# B&R Automation Studio project BrVideoPoker
Automation Studio 6.7.0.187; technology packages: mappServices 6.8.0, mappView 6.8.1, OpcUaCs 6.8.0

## Configuration Sim

CPU PC_any, AutomationRuntime D4.92, Build 11.3.0, Vc V4.72.5

### Task classes (Cpu.sw)
```
Cyclic#1:
  GameCode <- GameCode.prg
  UserSys <- UserSys.prg
  VisCtrl <- VisCtrl.prg
Binaries: arsvcreg, udbdef, TCData, arflatprv, arcoal, mvLoader, FWRules, Config_1, ashwac, User, sysconf, Config, asfw, arconfig, ashwd, Role, iomap
Libraries: PseudoRNG, AsIecCon, runtime, astime, AsIoTime, Cards, ArUser, arssl, ashw, arcert, fileio, sys_lib, aseth, dataobj, PokerHands, standard, MpUserX, MpBase
```

### Hardware
```
PC : PC_any v1.1.2.0 (OrderNumber=PC)
  ConfigurationID = BrVideoPoker_Sim
  FileDevice1
  FileDeviceName1 = USER
  FileDevicePath1 = USER_PATH
  ActivateOpcUa = 1
  OpcUa_SamplingTimer_Default = 4
  OpcUaInformationModels_PV_Version = 1
  ActivateFtpServer = 1
  ActivateWebServer = 1
  ActivateSdm = 1
```

### BRRole.brrole - PC/AccessAndSecurity/UserRoleSystem/BRRole.brrole
```
Element BR_Anonymous (Type=BRRole)
Element BR_Engineer (Type=BRRole)
Element BR_Observer (Type=BRRole)
Element BR_SafetyAdmin (Type=BRRole)
Element BR_SecurityAdmin (Type=BRRole)
```

- Physical/Sim/PC/IoMap.iom: same as Physical/Sim/PC/Cpu.per
- Physical/Sim/PC/PvMap.vvm: same as Physical/Sim/PC/Cpu.per
- Safety project (password-protected, skipped)

### Config.mpuserx - PC/mappServices/Config.mpuserx
```
Element UserMgmtX (Type=mpuserx)
  Mgr:
    AutoLogoutTime = 300
    UserNameLength = 3
    LoginAttempts = 5
  ServerSettings:
    Server:
      AdditionalUserData:
        [0] = mail
        [1] = telephoneNumber
  Groups:
    DefGroup#1:
      id = Administrators
      admin = TRUE
      rights:
        [0] = FullAccess
    DefGroup#2:
      id = Everyone
      level = 5
      admin = TRUE
```

### Config_1.mpuserxlogin - PC/mappServices/Config_1.mpuserxlogin
```
Element gUserXLogin (Type=mpuserxlogin)
```

## Configuration SuppC80

CPU 4PPC80.156B-13A, AutomationRuntime 6.8.1, Build 11.3.0

### Task classes (Cpu.sw)
```
Cyclic#1:
  GameCode <- GameCode.prg
  UserSys <- UserSys.prg
  VisCtrl <- VisCtrl.prg
Binaries: arsvcreg, udbdef, TCData, arflatprv, arcoal, mvLoader, FWRules, Config_1, ashwac, User, sysconf, Config, asfw, arconfig, ashwd, Role, iomap
Libraries: PseudoRNG, AsIecCon, runtime, astime, AsIoTime, Cards, ArUser, arssl, ashw, arcert, fileio, sys_lib, aseth, dataobj, PokerHands, standard, MpUserX, MpBase, AsBrStr
```

### Hardware
```
4PPC80_156B_13A : 4PPC80.156B-13A v1.4.0.0
  Connector IF2:
    AssignedOperatingSystem = ARemb
    ActivateDevice = 1
    ActivateSnmp = 2
  Connector IF3:
    OperatingSystem = ARemb
    ActivateDevice = 1
  Connector IF4:
    AssignedOperatingSystem = ARemb
  Connector IF5:
    AssignedOperatingSystem = GPOS
  Connector IF10:
    ActivateIna = 0
  ConfigurationID = BrVideoPoker_Sim
  Simulation = 1
  EnableDebugger = 1
  FileDevice1
  FileDeviceName1 = USER
  FileDevicePath1 = USER_PATH
  ActivateFtpServer = 1
  ActivateWebServer = 1
  ActivateSdm = 1
  LXTRemoteAccessUserWebGL = 
  LXTRemoteAccessPwdWebGL = 
```

- Physical/SuppC80/4PPC80_156B_13A/AccessAndSecurity/UserRoleSystem/BRRole.brrole: same as Physical/Sim/PC/AccessAndSecurity/UserRoleSystem/BRRole.brrole
- Physical/SuppC80/4PPC80_156B_13A/Cpu.per: same as Physical/Sim/PC/Cpu.per
- Physical/SuppC80/4PPC80_156B_13A/IoMap.iom: same as Physical/Sim/PC/Cpu.per
- Physical/SuppC80/4PPC80_156B_13A/PvMap.vvm: same as Physical/Sim/PC/Cpu.per
### Config.mpuserx - 4PPC80_156B_13A/mappServices/Config.mpuserx
```
Element UserMgmtX (Type=mpuserx)
  mapp.Gen:
    Audit = TRUE
  UserMgmtSystem:
    UserMgmtSystemType = 0
  ServerSettings:
    Server = ADServer
      Timeout = 10
      Mapping:
        TableName
      DisplayName = username
      AdditionalUserData:
        [0] = mail
        [1] = telephoneNumber
  PasswordPolicy:
    PasswordMaxAge = 0
    PasswordExpirationNotification = 0
    PasswordHistory = 0
    PasswordChangeReq = FALSE
    PasswordCase = TRUE
    PasswordAlpha = TRUE
    PasswordSpecial = TRUE
    PasswordLength = 8
  UserAccount:
    InvalidPasswordAttempts = 3
    UserExpirationTime = 0
    AutoLogoutTime = 3600
    UserNameLength = 1
    NoDelete = FALSE
    AdminUnlockTime = 3600
    EditSameLevel = 1
  ImportExport:
    ImportUser = 2
    ImportRole = 2
    ImportUnchecked = FALSE
    FileChecksum = 2
  Users:
    DefUser#1:
      id = Tester
      name
      lang
      measSystem = 0
  Roles:
    DefRole#1:
      id = Player
      level = 10
      admin = FALSE
```

- Physical/SuppC80/4PPC80_156B_13A/mappServices/Config_1.mpuserxlogin: same as Physical/Sim/PC/mappServices/Config_1.mpuserxlogin
## Logical view

Binary libraries used (declarations not repeated): operator, runtime, astime, AsIecCon, AsIoTime, ArUser, standard, MpUserX 6.8.0, MpBase 6.8.0, AsBrStr

### Global.typ - Global data types
```iecst
TYPE
	Player_typ : 	STRUCT
		Balance : REAL;
		Hand : ARRAY[0..4]OF Card_typ;
		HoldArr : ARRAY[0..4]OF BOOL;
		ChosenBet : REAL;
		Winnings : REAL;
		ActiveRound : BOOL;
		Result : FiveCardPoker_enum;
		LoggedIn : BOOL;
	END_STRUCT;
	Command_typ : 	STRUCT
		CMD_Confirm : BOOL;
		CMD_Action : BOOL;
	END_STRUCT;
END_TYPE
```

### Global.var - Global variables
```iecst
VAR
	gPlayer : Player_typ;
END_VAR
VAR CONSTANT
	BET_ARRAY : ARRAY[0..5] OF REAL := [0.1,0.2,0.5,1,2,5];
END_VAR
VAR
	gCurrentGame : GameVariant_enum;
	gCommand : Command_typ;
	gPayTable : PayTable_typ;
	gDeck : DeckFB;
	gPasswordInput : STRING[24];
	gUsernameInput : STRING[80];
END_VAR
```

### Package Logical/Libraries - Global libraries

### Library Logical/Libraries/Cards (IEC)

#### Types.typ - Exported data types
```iecst
TYPE
	Faces_enum :
		(
		CARD_TWO,
		CARD_THREE,
		CARD_FOUR,
		CARD_FIVE,
		CARD_SIX,
		CARD_SEVEN,
		CARD_EIGHT,
		CARD_NINE,
		CARD_TEN,
		CARD_JACK,
		CARD_QUEEN,
		CARD_KING,
		CARD_ACE
		);
	Suits_enum :
		(
		SUIT_HEARTS,
		SUIT_CLUBS,
		SUIT_DIAMONDS,
		SUIT_SPADES
		);
	Card_typ : 	STRUCT
		Face : Faces_enum;
		Suit : Suits_enum;
	END_STRUCT;
	DeckState :
		(
		DECKSTATE_INIT,
		DECKSTATE_IDLE,
		DECKSTATE_SHUFFLE,
		DECKSTATE_ERROR
		);
END_TYPE
```

#### Cards.fun - Exported functions and function blocks
```iecst
{REDUND_ERROR} FUNCTION SwapCard : BOOL (*Swap the place of two cards within deck*) (*$GROUP=User,$CAT=User,$GROUPICON=User.png,$CATICON=User.png*)
	VAR_INPUT
		Deck : REFERENCE TO ARRAY[0..51] OF Card_typ;
		CardIndexA : USINT;
		CardIndexB : USINT;
	END_VAR
	VAR
		TempCard : Card_typ;
	END_VAR
END_FUNCTION

FUNCTION_BLOCK DeckFB (*Core funciton block of the library*)
	VAR_INPUT
		CMD_Shuffle : BOOL;
		Enable : BOOL;
	END_VAR
	VAR_OUTPUT
		Deck : ARRAY[0..51] OF Card_typ;
		Active : BOOL;
		CommandDone : BOOL;
	END_VAR
	VAR
		IndexI : USINT;
		IndexJ : USINT;
		IndexR : USINT;
		ShuffleCount : USINT := 5;
		FaceIndex : USINT;
		SuitIndex : USINT;
		State : DeckState;
		Initialized : BOOL;
		Randy : PRNG;
	END_VAR
END_FUNCTION_BLOCK
```

#### CardsFB.st
```iecst
(* Deck Funtionality *)
FUNCTION_BLOCK DeckFB
	CASE State OF
		DECKSTATE_INIT:
			IF Enable AND NOT Initialized THEN
				//Initialize unshuffled deck
				FOR SuitIndex := 0 TO 3 DO
					FOR FaceIndex := 0 TO 12 DO
						Deck[SuitIndex*13+FaceIndex].Face := FaceIndex;
						Deck[SuitIndex*13+FaceIndex].Suit := SuitIndex;
					END_FOR;
				END_FOR;

				//Initialize RNG
				Randy(Multiplier := 4, Increment := 13, Seed := AsIOTimeStamp());

				State := DECKSTATE_IDLE;
				Active := TRUE;
				Initialized := TRUE;
			END_IF

		DECKSTATE_IDLE:
			IF CommandDone AND CMD_Shuffle THEN
				CommandDone := FALSE;
				CMD_Shuffle := FALSE;
			END_IF

			IF CMD_Shuffle THEN
				State := DECKSTATE_SHUFFLE;
			END_IF

		DECKSTATE_SHUFFLE:
			FOR IndexI := 0 TO ShuffleCount DO
				FOR IndexJ := 0 TO 51 DO
					Randy.CMD_Generate := TRUE;
					Randy();

					IndexR := UDINT_TO_USINT(  IndexJ + (Randy.Result MOD (52-IndexJ)));
					SwapCard(ADR(Deck), IndexJ, IndexR);
				END_FOR;
			END_FOR;

			CommandDone := TRUE;
			State := DECKSTATE_IDLE;

		DECKSTATE_ERROR:

	END_CASE;

END_FUNCTION_BLOCK
```

#### SwapCard.st
```iecst
(* Swap the place of two cards within deck *)
FUNCTION SwapCard
	TempCard := Deck[CardIndexA];
	Deck[CardIndexA] := Deck[CardIndexB];
	Deck[CardIndexB] := TempCard;
END_FUNCTION
```

### Library Logical/Libraries/PseudoRNG (IEC, version 1.00.1) - This library generates pseudo random numbers.

#### Constants.var - Exported constants
```iecst
VAR CONSTANT
	RAND_MAX : UINT := 32797; (*Maximum possible value for random number.*)
END_VAR
```

#### PseudoRNG.fun - Exported functions and function blocks
```iecst
FUNCTION_BLOCK PRNG
	VAR_INPUT
		Multiplier : {REDUND_UNREPLICABLE} UINT := 16; (*Multiplier parameter in formula*)
		Increment : {REDUND_UNREPLICABLE} UINT := 0; (*Increment parameter in formula*)
		CMD_Generate : {REDUND_UNREPLICABLE} BOOL; (*Input used to trigger generation*)
		Seed : UDINT; (*Initial seed used for formula*)
	END_VAR
	VAR_OUTPUT
		Result : {REDUND_UNREPLICABLE} UDINT; (*Output of generation*)
	END_VAR
	VAR
		Initialized : BOOL; (*True after procedure has been seeded*)
	END_VAR
END_FUNCTION_BLOCK
```

#### PRNG.st - Seeds and generates numbers using Linear Congruential Generation
```iecst
(* Psuedo Randon Number Generator *)
FUNCTION_BLOCK PRNG

	IF NOT Initialized THEN //Checks if prng has been seeded and does so if not
		Result := Seed; //Set initial "result" to the seed for purpose of the forumla
		Initialized := TRUE;
	END_IF

	IF CMD_Generate THEN //When CMD_Generate signal gets set to true generate the number
		Result := ((Result*Multiplier)+Increment) MOD RAND_MAX; //Formula applied to generate the next number
		CMD_Generate := FALSE; //Flips the trigger signal back false
	END_IF

END_FUNCTION_BLOCK
```

#### README.txt - PLEASE READ
```
Chris Hairston
chris.hairston@br-automation.com
4/1/2022

Overview:
	This library utilizes the linear congruential generator algorithm to generate a random number between 0 and 32797.

Linear Congruential Generation (LCG):
	NewNum = ((PrevNum*a) + c)% m
		where,
	a is the multiplier
	c is the increment
	m is the modulus (and functions as the max number, in this case 32767)

Usage:
	1. Seed the generator using AsIOTimeStamp
	2. Set CMD_Generate to true to generate number
	3. Call function block
	4. Use modulus function to determine range of prng (otherwise will be 0-32797)

Example: //This code generates a new number every 10 seconds.
	PROGRAM _INIT
		 Randy.Seed := DINT_TO_UDINT(AsIOTimeStamp());
	END_PROGRAM

	PROGRAM _CYCLIC
		TON_0(IN := NOT TON_0.Q, PT := T#10s);
		IF  TON_0.Q THEN
			Randy.CMD_Generate := TRUE;
		END_IF
		Randy();
		RandOf100 := Randy.Result MOD 100;
	END_PROGRAM
```

### Library Logical/Libraries/PokerHands (IEC)

#### Types.typ - Exported data types
```iecst
TYPE
	GameVariant_enum :
		(
		GAME_NONE,
		GAME_BONUS_POKER,
		GAME_DOUBLE_BONUS_POKER,
		GAME_TRIPLE_BONUS_POKER,
		GAME_ULTRA_BONUS_POKER,
		GAME_ALL_AMERICAN,
		GAME_JACKS_OR_BETTER,
		GAME_ACES_AND_EIGHTS,
		GAME_ACES_AND_FACES
		);
	FiveCardPoker_enum :
		(
		FIVECARDPOKER_NOTHING,
		FIVECARDPOKER_PAIR_FACE,
		FIVECARDPOKER_KINGS_OR_BETTER,
		FIVECARDPOKER_TWO_PAIR,
		FIVECARDPOKER_THREE_OF_A_KIND,
		FIVECARDPOKER_STRAIGHT,
		FIVECARDPOKER_FLUSH,
		FIVECARDPOKER_FULL_HOUSE,
		FIVECARDPOKER_FOUR_ANY,
		FIVECARDPOKER_FOUR_234,
		FIVECARDPOKER_FOUR_FIVE_THRU_K,
		FIVECARDPOKER_FOUR_SEVENS,
		FIVECARDPOKER_FOUR_EIGHTS,
		FIVECARDPOKER_FOUR_JQK,
		FIVECARDPOKER_FOUR_ACES,
		FIVECARDPOKER_STRAIGHT_FLUSH,
		FIVECARDPOKER_ROYAL_FLUSH
		);
	HandBools_typ : 	STRUCT
		AnyPair : BOOL;
		FacePair : BOOL;
		KingsOrBetter : BOOL;
		TwoPair : BOOL;
		ThreeOfAKind : BOOL;
		Straight : BOOL;
		Flush : BOOL;
		FourAny : BOOL;
		Four234 : BOOL;
		FourFiveThruKing : BOOL;
		FourSevens : BOOL;
		FourEights : BOOL;
		FourJQK : BOOL;
		FourAces : BOOL;
		Royal : BOOL;
	END_STRUCT;
	PayTable_typ : 	STRUCT
		Hands : ARRAY[0..13]OF FiveCardPoker_enum;
		WinningsScalarArr : ARRAY[0..13]OF REAL; (*Amount to multiply bet for winnings if that hand is achieved.*)
		GameVariant : GameVariant_enum;
	END_STRUCT;
	PayTableConst_typ : 	STRUCT
		Hands : ARRAY[0..13]OF USINT := [14(0)];
		WinningsScalarArr : ARRAY[0..13]OF REAL; (*Amount to multiply bet for winnings if that hand is achieved.*)
		GameVariant : USINT;
	END_STRUCT;
END_TYPE
```

#### Constants.var - Exported constants
```iecst
VAR CONSTANT
	PAY_TABLE_JACKS_OR_BETTER : PayTable_typ := (Hands:=[FIVECARDPOKER_ROYAL_FLUSH,FIVECARDPOKER_STRAIGHT_FLUSH,FIVECARDPOKER_FOUR_ANY,FIVECARDPOKER_FULL_HOUSE,FIVECARDPOKER_FLUSH,FIVECARDPOKER_STRAIGHT,FIVECARDPOKER_THREE_OF_A_KIND,FIVECARDPOKER_TWO_PAIR,FIVECARDPOKER_PAIR_FACE,FIVECARDPOKER_NOTHING,4(0)],WinningsScalarArr:=[250,50,25,9,6,4,3,2,1,5(0)],GameVariant:=GAME_JACKS_OR_BETTER); (*Pay Table for Jacks or Better*)
	PAY_TABLE_BONUS_POKER : PayTable_typ := (Hands:=[FIVECARDPOKER_ROYAL_FLUSH,FIVECARDPOKER_STRAIGHT_FLUSH,FIVECARDPOKER_FOUR_ACES,FIVECARDPOKER_FOUR_234,FIVECARDPOKER_FOUR_ANY,FIVECARDPOKER_FULL_HOUSE,FIVECARDPOKER_FLUSH,FIVECARDPOKER_STRAIGHT,FIVECARDPOKER_THREE_OF_A_KIND,FIVECARDPOKER_TWO_PAIR,FIVECARDPOKER_PAIR_FACE,3(0)],WinningsScalarArr:=[250,55,80,40,25,7,5,4,3,2,1,3(0.0)],GameVariant:=GAME_BONUS_POKER);
	PAY_TABLE_DOUBLE_BONUS_POKER : PayTable_typ := (Hands:=[FIVECARDPOKER_ROYAL_FLUSH,FIVECARDPOKER_STRAIGHT_FLUSH,FIVECARDPOKER_FOUR_ACES,FIVECARDPOKER_FOUR_234,FIVECARDPOKER_FOUR_ANY,FIVECARDPOKER_FULL_HOUSE,FIVECARDPOKER_FLUSH,FIVECARDPOKER_STRAIGHT,FIVECARDPOKER_THREE_OF_A_KIND,FIVECARDPOKER_TWO_PAIR,FIVECARDPOKER_PAIR_FACE,3(0)],WinningsScalarArr:=[250,50,160,80,50,10,7,5,3,2(1),3(0.0)],GameVariant:=GAME_DOUBLE_BONUS_POKER);
	PAY_TABLE_TRIPLE_BONUS_POKER : PayTable_typ := (Hands:=[FIVECARDPOKER_ROYAL_FLUSH,FIVECARDPOKER_STRAIGHT_FLUSH,FIVECARDPOKER_FOUR_ACES,FIVECARDPOKER_FOUR_234,FIVECARDPOKER_FOUR_ANY,FIVECARDPOKER_FULL_HOUSE,FIVECARDPOKER_FLUSH,FIVECARDPOKER_STRAIGHT,FIVECARDPOKER_THREE_OF_A_KIND,FIVECARDPOKER_TWO_PAIR,FIVECARDPOKER_KINGS_OR_BETTER,3(0)],WinningsScalarArr:=[250,50,240,120,75,9,7,4,3,2(1),3(0.0)],GameVariant:=GAME_TRIPLE_BONUS_POKER);
	PAY_TABLE_ULTRA_BONUS_POKER : PayTable_typ := (Hands:=[FIVECARDPOKER_ROYAL_FLUSH,FIVECARDPOKER_STRAIGHT_FLUSH,FIVECARDPOKER_FOUR_ACES,FIVECARDPOKER_FOUR_234,FIVECARDPOKER_FOUR_ANY,FIVECARDPOKER_FULL_HOUSE,FIVECARDPOKER_FLUSH,FIVECARDPOKER_STRAIGHT,FIVECARDPOKER_THREE_OF_A_KIND,FIVECARDPOKER_TWO_PAIR,FIVECARDPOKER_PAIR_FACE,3(0)],WinningsScalarArr:=[250,50,400,160,50,9,5,4,2,2(1),3(0.0)],GameVariant:=GAME_ULTRA_BONUS_POKER);
	PAY_TABLE_ALL_AMERICAN : PayTable_typ := (Hands:=[FIVECARDPOKER_ROYAL_FLUSH,FIVECARDPOKER_STRAIGHT_FLUSH,FIVECARDPOKER_FOUR_ANY,FIVECARDPOKER_FULL_HOUSE,FIVECARDPOKER_FLUSH,FIVECARDPOKER_STRAIGHT,FIVECARDPOKER_THREE_OF_A_KIND,FIVECARDPOKER_TWO_PAIR,FIVECARDPOKER_PAIR_FACE,FIVECARDPOKER_NOTHING,4(0)],WinningsScalarArr:=[800,200,30,3(8),3,2(1),5(0)],GameVariant:=GAME_ALL_AMERICAN);
	PAY_TABLE_ACES_AND_EIGHTS : PayTable_typ := (Hands:=[FIVECARDPOKER_ROYAL_FLUSH,FIVECARDPOKER_STRAIGHT_FLUSH,FIVECARDPOKER_FOUR_ACES,FIVECARDPOKER_FOUR_EIGHTS,FIVECARDPOKER_FOUR_SEVENS,FIVECARDPOKER_FOUR_ANY,FIVECARDPOKER_FULL_HOUSE,FIVECARDPOKER_FLUSH,FIVECARDPOKER_STRAIGHT,FIVECARDPOKER_THREE_OF_A_KIND,FIVECARDPOKER_TWO_PAIR,FIVECARDPOKER_PAIR_FACE,2(0)],WinningsScalarArr:=[250,50,2(80),50,25,8,5,4,3,2,1,2(0)],GameVariant:=GAME_ACES_AND_EIGHTS); (*Pay Table for Jacks or Better*)
	PAY_TABLE_ACES_AND_FACES : PayTable_typ := (Hands:=[FIVECARDPOKER_ROYAL_FLUSH,FIVECARDPOKER_STRAIGHT_FLUSH,FIVECARDPOKER_FOUR_ACES,FIVECARDPOKER_FOUR_JQK,FIVECARDPOKER_FOUR_ANY,FIVECARDPOKER_FULL_HOUSE,FIVECARDPOKER_FLUSH,FIVECARDPOKER_STRAIGHT,FIVECARDPOKER_THREE_OF_A_KIND,FIVECARDPOKER_TWO_PAIR,FIVECARDPOKER_PAIR_FACE,3(0)],WinningsScalarArr:=[500,50,80,40,25,8,5,4,3,2,1,3(0)],GameVariant:=GAME_ACES_AND_FACES); (*Pay Table for Jacks or Better*)
END_VAR
```

#### PokerHands.fun - Exported functions and function blocks
```iecst
{REDUND_ERROR} FUNCTION HandResult : FiveCardPoker_enum (*TODO: Add your comment here*) (*$GROUP=User,$CAT=User,$GROUPICON=User.png,$CATICON=User.png*)
	VAR_INPUT
		Hand : ARRAY[0..4] OF Card_typ;
		GameVariant : GameVariant_enum;
	END_VAR
	VAR
		ColumnTotals : ARRAY[1..14] OF USINT;
		RowTotals : ARRAY[0..3] OF USINT;
		i : USINT;
		j : USINT;
		k : USINT;
		CardMatrix : ARRAY[0..3,1..14] OF BOOL;
		tempHand : ARRAY[0..4] OF Card_typ;
		ResultBools : HandBools_typ;
		StraightCount : USINT;
		PairCount : USINT;
	END_VAR
END_FUNCTION

{REDUND_ERROR} FUNCTION CalculateWinnings : REAL (*TODO: Add your comment here*) (*$GROUP=User,$CAT=User,$GROUPICON=User.png,$CATICON=User.png*)
	VAR_INPUT
		PlayerHandResult : FiveCardPoker_enum;
		Bet : REAL;
	END_VAR
	VAR_IN_OUT
		PayTable : PayTable_typ;
	END_VAR
	VAR
		i : USINT;
	END_VAR
END_FUNCTION

FUNCTION Result2String : BOOL
	VAR_INPUT
		ResultHand : FiveCardPoker_enum;
	END_VAR
	VAR_IN_OUT
		destString : STRING[80];
	END_VAR
END_FUNCTION
```

#### CalculateWinnings.st
```iecst
(* TODO: Add your comment here *)
FUNCTION CalculateWinnings
	FOR i := 0 TO 13 DO
		IF PayTable.Hands[i] = PlayerHandResult THEN
			CalculateWinnings := Bet * PayTable.WinningsScalarArr[i];
			EXIT;
		END_IF
	END_FOR
END_FUNCTION
```

#### HandResult.st
```iecst
(* TODO: Add your comment here *)
FUNCTION HandResult
	//Initialization
	PairCount := 0;
	ResultBools.Royal := TRUE; //Will get turned false unless all cards "royal"
	//A matrix is used where there are 4 rows and 14 columns (Ace has a column for 1 and 14)
	//Because the card face enum starts with the 2 card at 0, we need to add 2
	FOR i := 0 TO 4 DO
		IF Hand[i].Face = CARD_ACE THEN
			CardMatrix[Hand[i].Suit,Hand[i].Face+2] := TRUE;
			CardMatrix[Hand[i].Suit,1] := TRUE;
		ELSE
			CardMatrix[Hand[i].Suit,Hand[i].Face+2] := TRUE;
		END_IF
	END_FOR

	FOR j := 0 TO 3 DO
		FOR k := 1 TO 14 DO
			IF CardMatrix[j,k] THEN

				IF k < 14 THEN //do not double count aces for the row total
					RowTotals[j] := RowTotals[j] + 1;
				END_IF

				ColumnTotals[k] := ColumnTotals[k] + 1;

			END_IF
		END_FOR
	END_FOR

	FOR j := 0 TO 3 DO //inspect the row totals
		IF RowTotals[j] = 5 THEN
			ResultBools.Flush := TRUE;
		END_IF
	END_FOR

	FOR k := 1 TO 14 DO //iterate through column totals
		IF ColumnTotals[k] = 4 THEN
			ResultBools.FourAny := TRUE;

			IF k = 8 THEN
				ResultBools.FourEights := TRUE;
			END_IF;

			IF k = 7 THEN
				ResultBools.FourSevens := TRUE;
			END_IF;

			IF k > 10 AND k < 14 THEN
				ResultBools.FourJQK := TRUE;
			END_IF

			IF k = 1 OR k = 14 THEN
				ResultBools.FourAces := TRUE;
			END_IF

			IF k >= 2 AND k <= 4 THEN
				ResultBools.Four234 := TRUE;
			END_IF

			IF k >=5 AND k <= 13 THEN
				ResultBools.FourFiveThruKing := TRUE;
			END_IF

		ELSIF ColumnTotals[k] = 3 THEN
			ResultBools.ThreeOfAKind := TRUE;

		ELSIF ColumnTotals[k] = 2 THEN
			IF k <> 1 THEN
				PairCount := PairCount + 1;
			END_IF

			ResultBools.AnyPair := TRUE;
			IF k >= 11 AND k <= 14 THEN
				ResultBools.FacePair := TRUE;
			END_IF

			IF k >= 12 AND k <= 14 THEN
				ResultBools.KingsOrBetter := TRUE;
			END_IF

		END_IF

		IF k >= 2 AND k<=9 AND ColumnTotals[k] > 0 THEN
			ResultBools.Royal := FALSE; //Fail royal check if any cards are not royal
		END_IF

		IF ColumnTotals[k] > 0 THEN
			StraightCount := StraightCount + 1;
			IF StraightCount = 5 THEN
				ResultBools.Straight := TRUE;
			END_IF
		ELSE
			StraightCount := 0;
		END_IF

	END_FOR

	IF PairCount >= 2 THEN
		ResultBools.TwoPair := TRUE;
	END_IF

	CASE GameVariant OF
		GAME_BONUS_POKER:
			//Large if statement based on hand result checks
			IF ResultBools.Royal AND ResultBools.Flush THEN
				HandResult := FIVECARDPOKER_ROYAL_FLUSH;
			ELSIF ResultBools.Straight AND ResultBools.Flush THEN
				HandResult := FIVECARDPOKER_STRAIGHT_FLUSH;
			ELSIF ResultBools.FourAces THEN
				HandResult := FIVECARDPOKER_FOUR_ACES;
			ELSIF ResultBools.Four234 THEN
				HandResult := FIVECARDPOKER_FOUR_234;
			ELSIF ResultBools.FourAny THEN
				HandResult := FIVECARDPOKER_FOUR_ANY;
			ELSIF ResultBools.ThreeOfAKind AND ResultBools.AnyPair THEN
				HandResult := FIVECARDPOKER_FULL_HOUSE;
			ELSIF ResultBools.Flush THEN
				HandResult := FIVECARDPOKER_FLUSH;
			ELSIF ResultBools.Straight THEN
				HandResult := FIVECARDPOKER_STRAIGHT;
			ELSIF ResultBools.ThreeOfAKind THEN
				HandResult := FIVECARDPOKER_THREE_OF_A_KIND;
			ELSIF ResultBools.TwoPair THEN
				HandResult := FIVECARDPOKER_TWO_PAIR;
			ELSIF ResultBools.FacePair THEN
				HandResult := FIVECARDPOKER_PAIR_FACE;
			ELSE
				HandResult := FIVECARDPOKER_NOTHING;
			END_IF

		GAME_DOUBLE_BONUS_POKER:
			//Large if statement based on hand result checks
			IF ResultBools.Royal AND ResultBools.Flush THEN
				HandResult := FIVECARDPOKER_ROYAL_FLUSH;
			ELSIF ResultBools.Straight AND ResultBools.Flush THEN
				HandResult := FIVECARDPOKER_STRAIGHT_FLUSH;
			ELSIF ResultBools.FourAces THEN
				HandResult := FIVECARDPOKER_FOUR_ACES;
			ELSIF ResultBools.Four234 THEN
				HandResult := FIVECARDPOKER_FOUR_234;
			ELSIF ResultBools.FourAny THEN
				HandResult := FIVECARDPOKER_FOUR_ANY;
			ELSIF ResultBools.ThreeOfAKind AND ResultBools.AnyPair THEN
				HandResult := FIVECARDPOKER_FULL_HOUSE;
			ELSIF ResultBools.Flush THEN
				HandResult := FIVECARDPOKER_FLUSH;
			ELSIF ResultBools.Straight THEN
				HandResult := FIVECARDPOKER_STRAIGHT;
			ELSIF ResultBools.ThreeOfAKind THEN
				HandResult := FIVECARDPOKER_THREE_OF_A_KIND;
			ELSIF ResultBools.TwoPair THEN
				HandResult := FIVECARDPOKER_TWO_PAIR;
			ELSIF ResultBools.FacePair THEN
				HandResult := FIVECARDPOKER_PAIR_FACE;
			ELSE
				HandResult := FIVECARDPOKER_NOTHING;
			END_IF

		GAME_TRIPLE_BONUS_POKER:
			//Large if statement based on hand result checks
			IF ResultBools.Royal AND ResultBools.Flush THEN
				HandResult := FIVECARDPOKER_ROYAL_FLUSH;
			ELSIF ResultBools.Straight AND ResultBools.Flush THEN
				HandResult := FIVECARDPOKER_STRAIGHT_FLUSH;
			ELSIF ResultBools.FourAces THEN
				HandResult := FIVECARDPOKER_FOUR_ACES;
			ELSIF ResultBools.Four234 THEN
				HandResult := FIVECARDPOKER_FOUR_234;
			ELSIF ResultBools.FourAny THEN
				HandResult := FIVECARDPOKER_FOUR_ANY;
			ELSIF ResultBools.ThreeOfAKind AND ResultBools.AnyPair THEN
				HandResult := FIVECARDPOKER_FULL_HOUSE;
			ELSIF ResultBools.Flush THEN
				HandResult := FIVECARDPOKER_FLUSH;
			ELSIF ResultBools.Straight THEN
				HandResult := FIVECARDPOKER_STRAIGHT;
			ELSIF ResultBools.ThreeOfAKind THEN
				HandResult := FIVECARDPOKER_THREE_OF_A_KIND;
			ELSIF ResultBools.TwoPair THEN
				HandResult := FIVECARDPOKER_TWO_PAIR;
			ELSIF ResultBools.KingsOrBetter THEN
				HandResult := FIVECARDPOKER_KINGS_OR_BETTER;
			ELSE
				HandResult := FIVECARDPOKER_NOTHING;
			END_IF
		GAME_ULTRA_BONUS_POKER:
			//Large if statement based on hand result checks
			IF ResultBools.Royal AND ResultBools.Flush THEN
				HandResult := FIVECARDPOKER_ROYAL_FLUSH;
			ELSIF ResultBools.Straight AND ResultBools.Flush THEN
				HandResult := FIVECARDPOKER_STRAIGHT_FLUSH;
			ELSIF ResultBools.FourAces THEN
				HandResult := FIVECARDPOKER_FOUR_ACES;
			ELSIF ResultBools.Four234 THEN
				HandResult := FIVECARDPOKER_FOUR_234;
			ELSIF ResultBools.FourAny THEN
				HandResult := FIVECARDPOKER_FOUR_ANY;
			ELSIF ResultBools.ThreeOfAKind AND ResultBools.AnyPair THEN
				HandResult := FIVECARDPOKER_FULL_HOUSE;
			ELSIF ResultBools.Flush THEN
				HandResult := FIVECARDPOKER_FLUSH;
			ELSIF ResultBools.Straight THEN
				HandResult := FIVECARDPOKER_STRAIGHT;
			ELSIF ResultBools.ThreeOfAKind THEN
				HandResult := FIVECARDPOKER_THREE_OF_A_KIND;
			ELSIF ResultBools.TwoPair THEN
				HandResult := FIVECARDPOKER_TWO_PAIR;
			ELSIF ResultBools.FacePair THEN
				HandResult := FIVECARDPOKER_PAIR_FACE;
			ELSE
				HandResult := FIVECARDPOKER_NOTHING;
			END_IF
		GAME_ALL_AMERICAN:
			//Large if statement based on hand result checks
			IF ResultBools.Royal AND ResultBools.Flush THEN
				HandResult := FIVECARDPOKER_ROYAL_FLUSH;
			ELSIF ResultBools.Straight AND ResultBools.Flush THEN
				HandResult := FIVECARDPOKER_STRAIGHT_FLUSH;
			ELSIF ResultBools.FourAny THEN
				HandResult := FIVECARDPOKER_FOUR_ANY;
			ELSIF ResultBools.ThreeOfAKind AND ResultBools.AnyPair THEN
				HandResult := FIVECARDPOKER_FULL_HOUSE;
			ELSIF ResultBools.Flush THEN
				HandResult := FIVECARDPOKER_FLUSH;
			ELSIF ResultBools.Straight THEN
				HandResult := FIVECARDPOKER_STRAIGHT;
			ELSIF ResultBools.ThreeOfAKind THEN
				HandResult := FIVECARDPOKER_THREE_OF_A_KIND;
			ELSIF ResultBools.TwoPair THEN
				HandResult := FIVECARDPOKER_TWO_PAIR;
			ELSIF ResultBools.FacePair THEN
				HandResult := FIVECARDPOKER_PAIR_FACE;
			ELSE
				HandResult := FIVECARDPOKER_NOTHING;
			END_IF
		GAME_JACKS_OR_BETTER:
			//Large if statement based on hand result checks
			IF ResultBools.Royal AND ResultBools.Flush THEN
				HandResult := FIVECARDPOKER_ROYAL_FLUSH;
			ELSIF ResultBools.Straight AND ResultBools.Flush THEN
				HandResult := FIVECARDPOKER_STRAIGHT_FLUSH;
			ELSIF ResultBools.FourAny THEN
				HandResult := FIVECARDPOKER_FOUR_ANY;
			ELSIF ResultBools.ThreeOfAKind AND ResultBools.AnyPair THEN
				HandResult := FIVECARDPOKER_FULL_HOUSE;
			ELSIF ResultBools.Flush THEN
				HandResult := FIVECARDPOKER_FLUSH;
			ELSIF ResultBools.Straight THEN
				HandResult := FIVECARDPOKER_STRAIGHT;
			ELSIF ResultBools.ThreeOfAKind THEN
				HandResult := FIVECARDPOKER_THREE_OF_A_KIND;
			ELSIF ResultBools.TwoPair THEN
				HandResult := FIVECARDPOKER_TWO_PAIR;
			ELSIF ResultBools.FacePair THEN
				HandResult := FIVECARDPOKER_PAIR_FACE;
			ELSE
				HandResult := FIVECARDPOKER_NOTHING;
			END_IF

		GAME_ACES_AND_EIGHTS:
			//Large if statement based on hand result checks
			IF ResultBools.Royal AND ResultBools.Flush THEN
				HandResult := FIVECARDPOKER_ROYAL_FLUSH;
			ELSIF ResultBools.Straight AND ResultBools.Flush THEN
				HandResult := FIVECARDPOKER_STRAIGHT_FLUSH;
			ELSIF ResultBools.FourAces THEN
				HandResult := FIVECARDPOKER_FOUR_ACES;
			ELSIF ResultBools.FourEights THEN
				HandResult := FIVECARDPOKER_FOUR_EIGHTS;
			ELSIF ResultBools.FourEights THEN
				HandResult := FIVECARDPOKER_FOUR_SEVENS;
			ELSIF ResultBools.FourAny THEN
				HandResult := FIVECARDPOKER_FOUR_ANY;
			ELSIF ResultBools.ThreeOfAKind AND ResultBools.AnyPair THEN
				HandResult := FIVECARDPOKER_FULL_HOUSE;
			ELSIF ResultBools.Flush THEN
				HandResult := FIVECARDPOKER_FLUSH;
			ELSIF ResultBools.Straight THEN
				HandResult := FIVECARDPOKER_STRAIGHT;
			ELSIF ResultBools.ThreeOfAKind THEN
				HandResult := FIVECARDPOKER_THREE_OF_A_KIND;
			ELSIF ResultBools.TwoPair THEN
				HandResult := FIVECARDPOKER_TWO_PAIR;
			ELSIF ResultBools.FacePair THEN
				HandResult := FIVECARDPOKER_PAIR_FACE;
			ELSE
				HandResult := FIVECARDPOKER_NOTHING;
			END_IF

		GAME_ACES_AND_FACES:
			//Large if statement based on hand result checks
			IF ResultBools.Royal AND ResultBools.Flush THEN
				HandResult := FIVECARDPOKER_ROYAL_FLUSH;
			ELSIF ResultBools.Straight AND ResultBools.Flush THEN
				HandResult := FIVECARDPOKER_STRAIGHT_FLUSH;
			ELSIF ResultBools.FourAces THEN
				HandResult := FIVECARDPOKER_FOUR_ACES;
			ELSIF ResultBools.FourJQK THEN
				HandResult := FIVECARDPOKER_FOUR_JQK;
			ELSIF ResultBools.FourAny THEN
				HandResult := FIVECARDPOKER_FOUR_ANY;
			ELSIF ResultBools.ThreeOfAKind AND ResultBools.AnyPair THEN
				HandResult := FIVECARDPOKER_FULL_HOUSE;
			ELSIF ResultBools.Flush THEN
				HandResult := FIVECARDPOKER_FLUSH;
			ELSIF ResultBools.Straight THEN
				HandResult := FIVECARDPOKER_STRAIGHT;
			ELSIF ResultBools.ThreeOfAKind THEN
				HandResult := FIVECARDPOKER_THREE_OF_A_KIND;
			ELSIF ResultBools.TwoPair THEN
				HandResult := FIVECARDPOKER_TWO_PAIR;
			ELSIF ResultBools.FacePair THEN
				HandResult := FIVECARDPOKER_PAIR_FACE;
			ELSE
				HandResult := FIVECARDPOKER_NOTHING;
			END_IF

	END_CASE
END_FUNCTION
```

#### Result2String.st
```iecst
FUNCTION Result2String
	CASE ResultHand OF
		FIVECARDPOKER_NOTHING:
			destString := '';
		FIVECARDPOKER_PAIR_FACE:
			destString := 'Jacks or Better';
		FIVECARDPOKER_KINGS_OR_BETTER:
			destString := 'Kings or Better';
		FIVECARDPOKER_TWO_PAIR:
			destString := 'Two Pair';
		FIVECARDPOKER_THREE_OF_A_KIND:
			destString := 'Three of a Kind';
		FIVECARDPOKER_FULL_HOUSE:
			destString := 'Full House';
		FIVECARDPOKER_STRAIGHT:
			destString := 'Straight';
		FIVECARDPOKER_FLUSH:
			destString := 'Flush';
		FIVECARDPOKER_STRAIGHT_FLUSH:
			destString := 'Straight Flush';
		FIVECARDPOKER_FOUR_ANY:
			destString := 'Four of a Kind';
		FIVECARDPOKER_FOUR_234:
			destString := 'Four 2s, 3s, 4s';
		FIVECARDPOKER_FOUR_FIVE_THRU_K:
			destString := 'Four 5s Thru Ks';
		FIVECARDPOKER_FOUR_SEVENS:
			destString := 'Four Sevens';
		FIVECARDPOKER_FOUR_EIGHTS:
			destString := 'Four Eights';
		FIVECARDPOKER_FOUR_JQK:
			destString := 'Four of a Face';
		FIVECARDPOKER_FOUR_ACES:
			destString := 'Four Aces';
		FIVECARDPOKER_ROYAL_FLUSH:
			destString := 'Royal Flush!';
	END_CASE;

	Result2String := TRUE; //Successful function call
END_FUNCTION
```

- Visualisation Logical/mappView (not shown)

### Program Logical/GameCode (IEC)

#### Main.st - Init, cyclic, exit code
```iecst
PROGRAM _INIT
	(* Insert code here *)
	 gCurrentGame;
END_PROGRAM

PROGRAM _CYCLIC
	 //TestTable := PAY_TABLE_JACKS_OR_BETTER;
	//gPlayer.Hand := TestHand;
	//Result := HandResult(gPlayer.Hand, GAME_JACKS_OR_BETTER);

	//Choose pay table based on game
	CASE gCurrentGame OF
		GAME_NONE:

		GAME_BONUS_POKER:
			gPayTable := PAY_TABLE_BONUS_POKER;
		GAME_DOUBLE_BONUS_POKER:
			gPayTable := PAY_TABLE_DOUBLE_BONUS_POKER;
		GAME_TRIPLE_BONUS_POKER:
			gPayTable := PAY_TABLE_TRIPLE_BONUS_POKER;
		GAME_ULTRA_BONUS_POKER:
			gPayTable := PAY_TABLE_ULTRA_BONUS_POKER;
		GAME_ALL_AMERICAN:
			gPayTable := PAY_TABLE_ALL_AMERICAN;
		GAME_JACKS_OR_BETTER:
			gPayTable := PAY_TABLE_JACKS_OR_BETTER;
		GAME_ACES_AND_EIGHTS:
			gPayTable := PAY_TABLE_ACES_AND_EIGHTS;
		GAME_ACES_AND_FACES:
			gPayTable := PAY_TABLE_ACES_AND_FACES;
	END_CASE

	CASE GameState OF
		GAME_STATE_WAIT:
			gPlayer.Result := FIVECARDPOKER_NOTHING;
			gPlayer.Winnings := 0;
			gPlayer.ActiveRound := FALSE;

			ActionButtonStr := 'Play';

			IF gCommand.CMD_Action THEN
				gCommand.CMD_Action := FALSE;
				GameState := GAME_STATE_SHUFFLE;
			END_IF

		GAME_STATE_SHUFFLE:
			gDeck.CMD_Shuffle := TRUE;

			IF gDeck.CommandDone THEN
				GameState := GAME_STATE_DEAL;
			END_IF

		GAME_STATE_DEAL:
			gPlayer.ActiveRound := TRUE;
			gPlayer.Balance := gPlayer.Balance - gPlayer.ChosenBet;
			FOR DeckCardCount := 0 TO 4 DO
				gPlayer.Hand[DeckCardCount] := gDeck.Deck[DeckCardCount];
			END_FOR

			GameState := GAME_STATE_HOLD;

		GAME_STATE_HOLD:
			//Wait for user to select cards to hold
			ActionButtonStr := 'Draw';
			IF NOT gPlayer.LoggedIn THEN
				GameState := GAME_STATE_WAIT;
			ELSIF gCommand.CMD_Action THEN
				gCommand.CMD_Action := FALSE;
				GameState := GAME_STATE_REDEAL;
			END_IF

		GAME_STATE_REDEAL:
			DeckCardCount := 5;

			FOR i := 0 TO 4 DO
				IF  NOT gPlayer.HoldArr[i] THEN
					gPlayer.Hand[i] := gDeck.Deck[DeckCardCount];
					DeckCardCount := DeckCardCount + 1;
				ELSE
					gPlayer.HoldArr[i] := FALSE;
				END_IF
			END_FOR

			GameState := GAME_STATE_RESULTS;

		GAME_STATE_RESULTS:
			gPlayer.Result := HandResult(gPlayer.Hand, gCurrentGame);
			ActionButtonStr := 'Clear';

			gPlayer.Winnings := CalculateWinnings(gPlayer.Result, gPlayer.ChosenBet, gPayTable);

			IF R_TRIG_ResultState.Q THEN
				gPlayer.Balance := gPlayer.Balance + gPlayer.Winnings;
			END_IF

			IF NOT gPlayer.LoggedIn THEN
				GameState := GAME_STATE_WAIT;
			ELSIF gCommand.CMD_Confirm OR gCommand.CMD_Action THEN
				gCommand.CMD_Action := FALSE;
				gCommand.CMD_Confirm := FALSE;
				GameState := GAME_STATE_WAIT;
			END_IF

		GAME_STATE_ERROR:

	END_CASE

	//R Trig to ensure winnings are only given once
	R_TRIG_ResultState(CLK := (GameState = GAME_STATE_RESULTS));

	//Deck custom FB
	gDeck.Enable := TRUE;
	gDeck();

END_PROGRAM

PROGRAM _EXIT
	(* Insert code here *)

END_PROGRAM
```

#### Types.typ - Local data types
```iecst
TYPE
	GameState_enum :
		(
		GAME_STATE_WAIT,
		GAME_STATE_SHUFFLE,
		GAME_STATE_DEAL,
		GAME_STATE_HOLD,
		GAME_STATE_REDEAL,
		GAME_STATE_RESULTS,
		GAME_STATE_ERROR
		);
END_TYPE
```

#### Variables.var - Local variables
```iecst
VAR
	TestHand : ARRAY[0..4] OF Card_typ := [(Face:=CARD_ACE,Suit:=SUIT_HEARTS),(Face:=CARD_TWO,Suit:=SUIT_CLUBS),(Face:=CARD_THREE,Suit:=SUIT_DIAMONDS),(Face:=CARD_FOUR,Suit:=SUIT_SPADES),(Face:=CARD_FIVE,Suit:=SUIT_HEARTS)];
	GameState : GameState_enum;
	DeckCardCount : USINT;
	i : USINT;
	R_TRIG_ResultState : R_TRIG;
	ActionButtonStr : STRING[80];
END_VAR
```

### Program Logical/UserSys (IEC)

#### Main.st - Init, cyclic, exit code
```iecst
PROGRAM _INIT

END_PROGRAM

PROGRAM _CYCLIC
	CASE UserState OF
		USERSTATE_WAITINGFORUSER:
			gPlayer.Balance := 0;
			ArUserSetProperty_FB.Execute := FALSE;
			gPlayer.LoggedIn := FALSE;

			IF CurrentUser <> '' AND CurrentUser <> 'Anonymous' THEN
				UserState := USERSTATE_GETBALANCE;
			END_IF;

		USERSTATE_GETBALANCE:
			ArUserGetProperty_FB.ElementName := CurrentUser;
			ArUserGetProperty_FB.ElementType := arUSER_USER_PROPERTIES;
			ArUserGetProperty_FB.PropertyName := 'Balance';
			ArUserGetProperty_FB.Execute := TRUE;

			gPlayer.LoggedIn := TRUE;

			//-1070585892: Specified element does not exist
			IF ArUserGetProperty_FB.Error AND ArUserGetProperty_FB.ErrorID = arUSER_ERR_DOES_NOT_EXIST THEN //if property doesnt exist we will create it
				UserState := USERSTATE_RUN;
				gPlayer.Balance := 100;
				ArUserGetProperty_FB.Execute := FALSE;
			ELSIF ArUserGetProperty_FB.Done THEN
				UserState := USERSTATE_RUN;
				gPlayer.Balance := STRING_TO_REAL(ArUserGetProperty_FB.PropertyValue);
				ArUserGetProperty_FB.Execute := FALSE;
			ELSIF ArUserGetProperty_FB.Error THEN
				UserState := USERSTATE_ERROR;
				ArUserGetProperty_FB.Execute := FALSE;
			END_IF

		USERSTATE_RUN:
			//ArUserSetProperty_0(Execute := , ElementType := , ElementName := , PropertyName := , PropertyValue := );
			ArUserSetProperty_FB.ElementName := CurrentUser;
			ArUserSetProperty_FB.ElementType := arUSER_USER_PROPERTIES;
			ArUserSetProperty_FB.PropertyName := 'Balance';
			ArUserSetProperty_FB.PropertyValue := REAL_TO_STRING(gPlayer.Balance);
			ArUserSetProperty_FB.Execute := TRUE;

			IF ArUserSetProperty_FB.Done THEN
				ArUserSetProperty_FB.Execute := FALSE;
			END_IF

			IF CurrentUser = '' OR CurrentUser = 'Anonymous' THEN
				UserState := USERSTATE_WAITINGFORUSER;
				ArUserSetProperty_FB.Execute := FALSE;
			END_IF;

		USERSTATE_ERROR:

	END_CASE;

	CASE CreateUserState OF
		CREATE_USER_WAIT:
			IF CMD_CreateUser THEN
				CreateUserState := CREATE_USER_CREATE;
				//CMD_UserCreationDone := FALSE;
			END_IF

		CREATE_USER_CREATE:
			ArUserCreate_FB.Execute := TRUE;
			ArUserCreate_FB.UserName := gUsernameInput;

			IF ArUserCreate_FB.Busy THEN
				//do nothing
			ELSIF ArUserCreate_FB.Error THEN
				ArUserCreate_FB.Execute := FALSE;
				ArUserCreate_FB.UserName := '';
				ErrorCode := ArUserCreate_FB.ErrorID;
				CreateUserState := CREATE_USER_ERROR;
			ELSIF ArUserCreate_FB.Done THEN
				//CMD_CreateUser := FALSE;
				ArUserCreate_FB.Execute := FALSE;
				ArUserCreate_FB.UserName := '';
				CreateUserState := CREATE_USER_SET_PASSWORD;
			END_IF

		CREATE_USER_SET_PASSWORD:
			ArUserSetPassword_FB.Execute := TRUE;
			ArUserSetPassword_FB.UserName := gUsernameInput;
			ArUserSetPassword_FB.Password := gPasswordInput;

			IF ArUserSetPassword_FB.Busy THEN
				//do nothing
			ELSIF ArUserSetPassword_FB.Error THEN
				ArUserSetPassword_FB.Execute := FALSE;
				ArUserSetPassword_FB.UserName := '';
				ArUserSetPassword_FB.Password := '';
				ErrorCode := ArUserSetPassword_FB.ErrorID;
				CreateUserState := CREATE_USER_ERROR;
			ELSIF ArUserSetPassword_FB.Done THEN
				//CMD_CreateUser := FALSE;
				ArUserSetPassword_FB.Execute := FALSE;
				ArUserSetPassword_FB.UserName := '';
				ArUserSetPassword_FB.Password := '';
				CreateUserState := CREATE_USER_ASSIGN_ROLE;
			END_IF

		CREATE_USER_ASSIGN_ROLE:
			ArUserAssignRole_FB.Execute := TRUE;
			ArUserAssignRole_FB.UserName := gUsernameInput;
			ArUserAssignRole_FB.RoleName := 'Player';
			IF ArUserAssignRole_FB.Busy THEN
				//do nothing
			ELSIF ArUserAssignRole_FB.Error THEN
				ArUserAssignRole_FB.Execute := FALSE;
				ArUserAssignRole_FB.UserName := '';
				ArUserAssignRole_FB.RoleName := '';
				ErrorCode := ArUserAssignRole_FB.ErrorID;
				CreateUserState := CREATE_USER_ERROR;
			ELSIF ArUserAssignRole_FB.Done THEN
				ArUserAssignRole_FB.Execute := FALSE;
				ArUserAssignRole_FB.UserName := '';
				ArUserAssignRole_FB.RoleName := '';
				ErrorCode := 0;
				ErrorStr := '';
				CMD_UserCreationDone := TRUE;
				CMD_CreateUser := FALSE;
				CreateUserState := CREATE_USER_WAIT; //go to user state, if no error it will progress to wait
			END_IF

		CREATE_USER_ERROR:
			CMD_CreateUser := FALSE;
			CreateUserState := CREATE_USER_WAIT;
			CASE ErrorCode OF
				arUSER_ERR_PARAMETER:
					ErrorStr := 'The function block was called with an invalid parameter.'; //Should not occur unless programmer has messed up
				arUSER_ERR_ALREADY_EXISTS:
					ErrorStr := 'The user already exists.';
				arUSER_ERR_DOES_NOT_EXIST:
					ErrorStr := 'The user does not exist.';
				arUSER_ERR_INTERNAL:
					ErrorStr :='An unexpected internal error has occurred.';
				ELSE
					ErrorStr := 'An unspecified error has occured. Check the logger.';
			END_CASE

	END_CASE

	ArUserCreate_FB();
	ArUserSetPassword_FB();
	ArUserGetProperty_FB();
	ArUserSetProperty_FB();
	ArUserAssignRole_FB();

	//MpUserXManagerUI for monitoring (requres mpuserxlogin)
	MpUserXLogin_FB(MpLink :=  ADR(gUserXLogin), Enable := TRUE);
	MpUserXManagerUI_FB(MpLink := ADR(gUserXLogin), Enable := TRUE, UISetup := MpUserXManagerUI_Setup, UIConnect := ADR(MpUserXManagerUI_Connect));
END_PROGRAM

PROGRAM _EXIT
	(* Insert code here *)

END_PROGRAM
```

#### Types.typ - Local data types
```iecst
TYPE
	UserState_enum :
		(
		USERSTATE_WAITINGFORUSER,
		USERSTATE_GETBALANCE,
		USERSTATE_RUN,
		USERSTATE_LOGOUT,
		USERSTATE_ERROR
		);
	CreateUserState_enum :
		(
		CREATE_USER_WAIT,
		CREATE_USER_CREATE,
		CREATE_USER_SET_PASSWORD,
		CREATE_USER_ASSIGN_ROLE,
		CREATE_USER_HMI_ACKNOWLEDGE,
		CREATE_USER_ERROR
		);
END_TYPE
```

#### Variables.var - Local variables
```iecst
VAR
	CMD_UserCreationAcknowledged : USINT;
	CMD_CreateUser : BOOL;
	CurrentUser : STRING[80];
	ArUserSetProperty_FB : ArUserSetProperty;
	CreateUserPassStr : STRING[80];
	CreateUserNameStr : STRING[80];
	ArUserCreate_FB : ArUserCreate;
	ArUserSetPassword_FB : ArUserSetPassword;
	ArUserGetProperty_FB : ArUserGetProperty;
	UserState : UserState_enum;
	MpUserXManagerUI_Connect : MpUserXMgrUIConnectType;
	MpUserXManagerUI_Setup : MpUserXMgrUISetupType;
	MpUserXLogin_FB : MpUserXLogin;
	MpUserXManagerUI_FB : MpUserXManagerUI;
	CreateUserState : CreateUserState_enum;
	ErrorCode : DINT;
	ErrorStr : STRING[80];
	CMD_UserCreationDone : BOOL;
	ArUserAssignRole_FB : ArUserAssignRole;
END_VAR
```

### Program Logical/VisCtrl (IEC)

#### Main.st - Init, cyclic, exit code
```iecst
PROGRAM _INIT
	(* Insert code here *)

END_PROGRAM

PROGRAM _CYCLIC
	(* Insert code here *)
	//ensure password input meets requirements and if so enable the confirm button for user creation

	//transfer the string to an ascii array
	brsmemcpy(ADR(pwAsciiArray), ADR(gPasswordInput), brsstrlen(ADR(gPasswordInput)));

	//Reset values before restarting loop
	pwReqCheck := pwReqCheck_NULL;

	//Ensure password is at least 8 characters long
	pwReqCheck.isMinLength := brsstrlen(ADR(gPasswordInput)) >= 8;

	FOR pwReqCheckIndex := 0 TO brsstrlen(ADR(gPasswordInput)) DO //loop through full pw string
		//check for upper and lower case
		IF pwAsciiArray[pwReqCheckIndex] >= 65 AND pwAsciiArray[pwReqCheckIndex] <= 90 THEN
			pwReqCheck.hasUpperCase := TRUE;
		ELSIF pwAsciiArray[pwReqCheckIndex] >= 97 AND pwAsciiArray[pwReqCheckIndex] <= 122 THEN
			pwReqCheck.hasLowerCase := TRUE;
		END_IF

		//check for alphanumeric characters
		IF (pwAsciiArray[pwReqCheckIndex] >= 48 AND pwAsciiArray[pwReqCheckIndex] <= 57) OR (pwAsciiArray[pwReqCheckIndex] >= 65 AND pwAsciiArray[pwReqCheckIndex] <= 90) OR (pwAsciiArray[pwReqCheckIndex] >= 97 AND pwAsciiArray[pwReqCheckIndex] <= 122) THEN
			pwReqCheck.hasAlphaNumericChars := TRUE;
		END_IF

		//check for special characters
		IF (pwAsciiArray[pwReqCheckIndex] >= 33 AND pwAsciiArray[pwReqCheckIndex] <= 47) OR (pwAsciiArray[pwReqCheckIndex] >= 58 AND pwAsciiArray[pwReqCheckIndex] <= 64) OR (pwAsciiArray[pwReqCheckIndex] >= 123 AND pwAsciiArray[pwReqCheckIndex] <= 126) THEN
			pwReqCheck.hasSpecialChars := TRUE;
		END_IF
	END_FOR;

	//if lower and upper case letters are found during the loop then the pw is mixed case
	pwReqCheck.isMixedCase := pwReqCheck.hasLowerCase AND pwReqCheck.hasUpperCase;

	//if all requirements are met, the confirmation button is enabled
	enableCreateUser := pwReqCheck.isMinLength AND pwReqCheck.isMixedCase AND pwReqCheck.hasAlphaNumericChars AND pwReqCheck.hasSpecialChars;

	gPlayer.ChosenBet := BET_ARRAY[BetIndex];

	//Generate card strings for the image bindings
	FOR i :=0 TO 4 DO
		IF NOT gPlayer.ActiveRound THEN
			CardStr[i] := 	'Media/Cards/Minicard_Back.svg';
		ELSE
			CardStr[i] := 'Media/Cards/Minicard_';

			//CASE statement for card value/face
			CASE gPlayer.Hand[i].Face OF
				CARD_TWO:
					CardStr[i] := CONCAT(CardStr[i], '2');
				CARD_THREE:
					CardStr[i] := CONCAT(CardStr[i], '3');
				CARD_FOUR:
					CardStr[i] := CONCAT(CardStr[i], '4');
				CARD_FIVE:
					CardStr[i] := CONCAT(CardStr[i], '5');
				CARD_SIX:
					CardStr[i] := CONCAT(CardStr[i], '6');
				CARD_SEVEN:
					CardStr[i] := CONCAT(CardStr[i], '7');
				CARD_EIGHT:
					CardStr[i] := CONCAT(CardStr[i], '8');
				CARD_NINE:
					CardStr[i] := CONCAT(CardStr[i], '9');
				CARD_TEN:
					CardStr[i] := CONCAT(CardStr[i], '10');
				CARD_JACK:
					CardStr[i] := CONCAT(CardStr[i], 'J');
				CARD_QUEEN:
					CardStr[i] := CONCAT(CardStr[i], 'Q');
				CARD_KING:
					CardStr[i] := CONCAT(CardStr[i], 'K');
				CARD_ACE:
					CardStr[i] := CONCAT(CardStr[i], 'A');
			END_CASE

			CASE gPlayer.Hand[i].Suit OF
				SUIT_CLUBS:
					CardStr[i] := CONCAT(CardStr[i], 'C');
				SUIT_DIAMONDS:
					CardStr[i] := CONCAT(CardStr[i], 'D');
				SUIT_HEARTS:
					CardStr[i] := CONCAT(CardStr[i], 'H');
				SUIT_SPADES:
					CardStr[i] := CONCAT(CardStr[i], 'S');
			END_CASE

			CardStr[i] := CONCAT(CardStr[i], '.svg');
		END_IF
	END_FOR

	Result2String(gPlayer.Result, ResultStr);

	CASE gCurrentGame OF
		GAME_NONE:
			GameStr := '';
		GAME_BONUS_POKER:
			GameStr := 'Bonus Poker';
		GAME_DOUBLE_BONUS_POKER:
			GameStr := 'Double Bonus Poker';
		GAME_TRIPLE_BONUS_POKER:
			GameStr := 'Triple Bonus Poker';
		GAME_ULTRA_BONUS_POKER:
			GameStr := 'Ultra Bonus Poker';
		GAME_ALL_AMERICAN:
			GameStr := 'All American';
		GAME_JACKS_OR_BETTER:
			GameStr := 'Jacks or Better';
		GAME_ACES_AND_EIGHTS:
			GameStr := 'Aces & Eights';
		GAME_ACES_AND_FACES:
			GameStr := 'Aces & Faces';
	END_CASE

	EnableBetting := NOT gPlayer.ActiveRound; //Betting should only be enabled when the round is not active
	NotLoggedIn := NOT gPlayer.LoggedIn;

	FOR i := 0 TO 13 DO
		Result2String(gPayTable.Hands[i], PayTableStr[i]);
		PayTableScaledWinnings[i] := gPayTable.WinningsScalarArr[i] * gPlayer.ChosenBet;
		PayTableVisible[i] := gPayTable.WinningsScalarArr[i] <> 0;
	END_FOR

END_PROGRAM

PROGRAM _EXIT
	(* Insert code here *)

END_PROGRAM
```

#### Types.typ - Local data types
```iecst
TYPE
	pwReqCheck_typ : 	STRUCT
		isMixedCase : BOOL;
		isMinLength : BOOL;
		hasSpecialChars : BOOL;
		hasAlphaNumericChars : BOOL;
		hasLowerCase : BOOL;
		hasUpperCase : BOOL;
	END_STRUCT;
END_TYPE
```

#### Variables.var - Local variables
```iecst
VAR
	enableCreateUser : BOOL;
END_VAR
VAR CONSTANT
	pwReqCheck_NULL : pwReqCheck_typ := (0);
END_VAR
VAR
	pwReqCheck : pwReqCheck_typ;
	pwInput : STRING[80];
	CardStr : ARRAY[0..4] OF STRING[80];
	BetIndex : USINT;
	i : USINT;
	ResultStr : STRING[80];
	EnableBetting : BOOL;
	GameStr : STRING[80];
	NotLoggedIn : BOOL;
	PayTableStr : ARRAY[0..13] OF STRING[80];
	PayTableScaledWinnings : ARRAY[0..13] OF REAL;
	PayTableVisible : ARRAY[0..13] OF BOOL;
	pwReqCheckIndex : UDINT;
	pwAsciiArray : ARRAY[0..23] OF USINT;
END_VAR
```
